(* IEC 61131-3 sources: iec-st-tools/testdata/src/UserTypes, 1 file *)

(* ---- TestTypes.st ---- *)
TYPE
    TestStruct : STRUCT
        Value   : INT := 0;
        IsValid : BOOL := FALSE;
        Name    : STRING := '';
    END_STRUCT;

    TestEnum : (
        stIdle   := 0,
        stactive := 1,
        stError  := 2
    );
END_TYPE
